(* IEC 61131-3 sources: nautilus/website/lessons/b1-blink/variants/ok-restart-by-reset, 1 file *)

(* ---- program.st ---- *)
PROGRAM Blink
VAR
    tick : TON;
    flip : BOOL;
END_VAR
tick(IN := NOT flip, PT := T#500ms);
flip := tick.Q;
IF flip THEN
    Lamp := NOT Lamp;
END_IF;
END_PROGRAM
